Staubli VAL3: utData.pjx

--- utData.pjx ---
Parameters version=s8.8.3Cs9_BS1660 stackSize=5000 millimeterUnit=true
Program file=start.pgx
Program file=stop.pgx
Data file=utData.dtx

--- utData.dtx ---
public num nVal
public bool bStatus

--- start.pgx ---
program start()
begin
end

--- stop.pgx ---
program stop()
begin
end
